Fanuc KAREL source: KO00116.KL

PROGRAM KO00116
%NOLOCKGROUP
VAR
  A: ARRAY[2] OF BYTE
  B: REAL
  OUT: REAL
BEGIN
  A[1] = 1
  B = 2
  OUT = ATAN2(A[1], B)
END KO00116
